// Mitsubishi GX Works2 project: TEAM_PLC   PLC: Q03UD

PROGRAM MAIN3
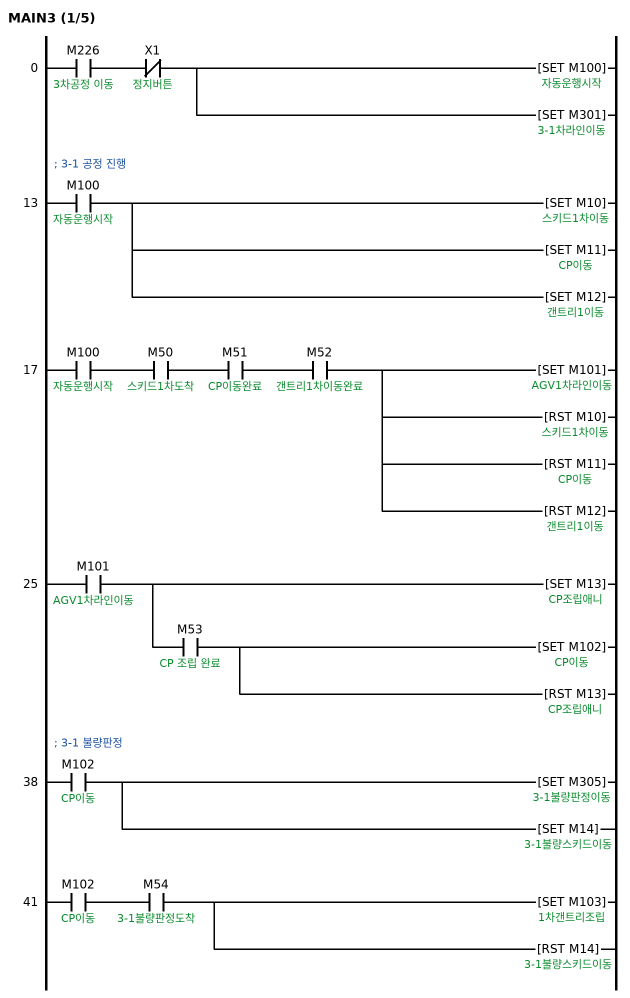
0     LD      M226  ; 3차공정 이동
      ANI     X1  ; 정지버튼
      SET     M100  ; 자동운행시작
      SET     M301  ; 3-1차라인이동
; 3-1 공정 진행
13    LD      M100  ; 자동운행시작
      SET     M10  ; 스키드1차이동
      SET     M11  ; CP이동
      SET     M12  ; 갠트리1이동
17    LD      M100  ; 자동운행시작
      AND     M50  ; 스키드1차도착
      AND     M51  ; CP이동완료
      AND     M52  ; 갠트리1차이동완료
      SET     M101  ; AGV1차라인이동
      RST     M10  ; 스키드1차이동
      RST     M11  ; CP이동
      RST     M12  ; 갠트리1이동
25    LD      M101  ; AGV1차라인이동
      SET     M13  ; CP조립애니
      AND     M53  ; CP 조립 완료
      SET     M102  ; CP이동
      RST     M13  ; CP조립애니
; 3-1 불량판정
38    LD      M102  ; CP이동
      SET     M305  ; 3-1불량판정이동
      SET     M14  ; 3-1불량스키드이동
41    LD      M102  ; CP이동
      AND     M54  ; 3-1불량판정도착
      SET     M103  ; 1차갠트리조립
      RST     M14  ; 3-1불량스키드이동
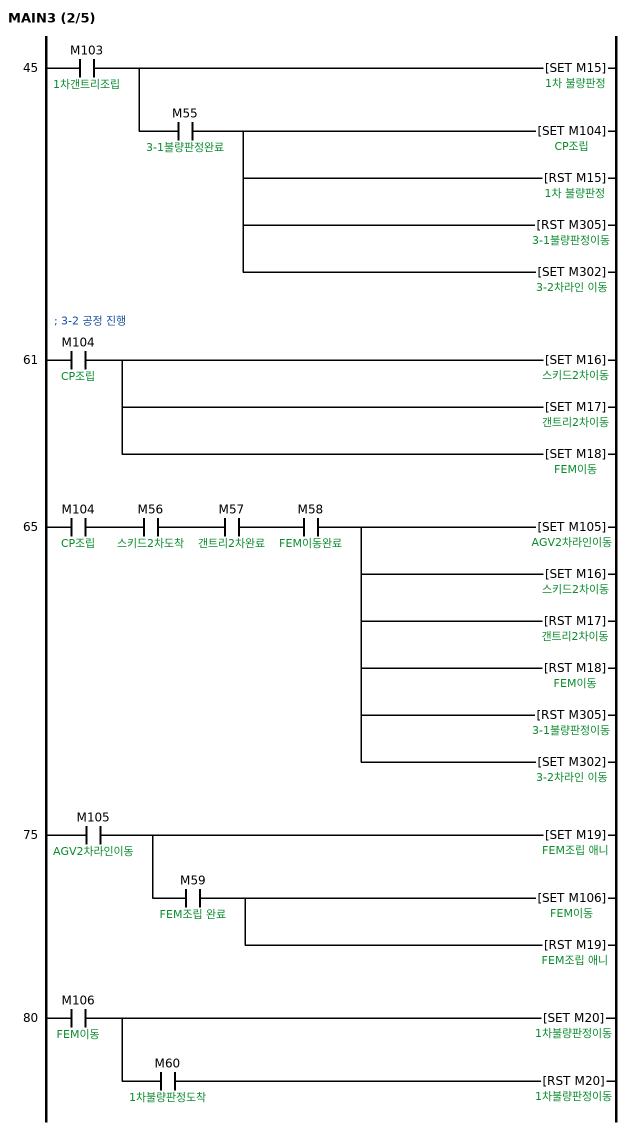
45    LD      M103  ; 1차갠트리조립
      SET     M15  ; 1차 불량판정
      AND     M55  ; 3-1불량판정완료
      SET     M104  ; CP조립
      RST     M15  ; 1차 불량판정
      RST     M305  ; 3-1불량판정이동
      SET     M302  ; 3-2차라인 이동
; 3-2 공정 진행
61    LD      M104  ; CP조립
      SET     M16  ; 스키드2차이동
      SET     M17  ; 갠트리2차이동
      SET     M18  ; FEM이동
65    LD      M104  ; CP조립
      AND     M56  ; 스키드2차도착
      AND     M57  ; 갠트리2차완료
      AND     M58  ; FEM이동완료
      SET     M105  ; AGV2차라인이동
      SET     M16  ; 스키드2차이동
      RST     M17  ; 갠트리2차이동
      RST     M18  ; FEM이동
      RST     M305  ; 3-1불량판정이동
      SET     M302  ; 3-2차라인 이동
75    LD      M105  ; AGV2차라인이동
      SET     M19  ; FEM조립 애니
      AND     M59  ; FEM조립 완료
      SET     M106  ; FEM이동
      RST     M19  ; FEM조립 애니
80    LD      M106  ; FEM이동
      SET     M20  ; 1차불량판정이동
      AND     M60  ; 1차불량판정도착
      RST     M20  ; 1차불량판정이동
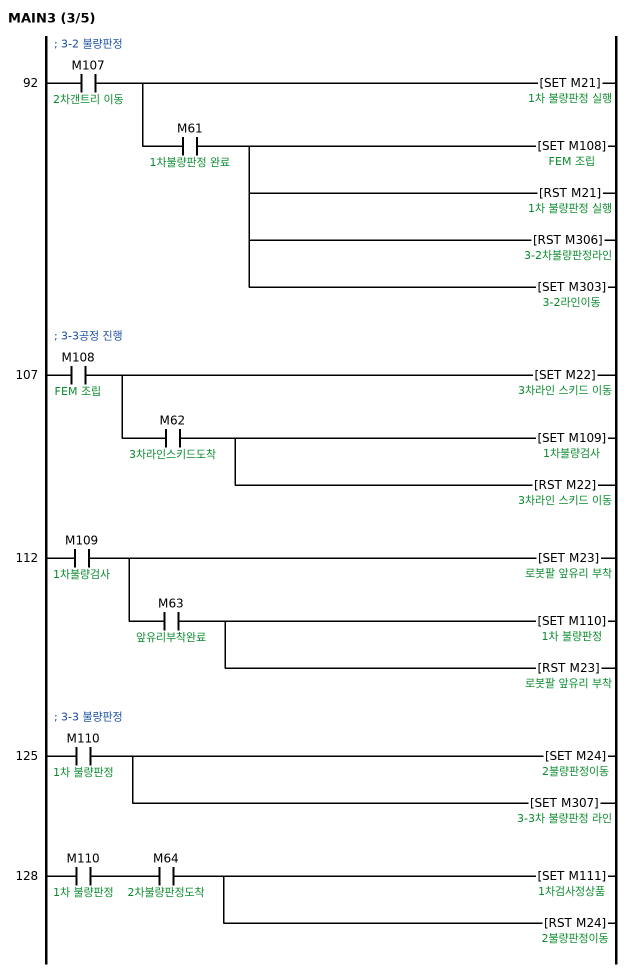
; 3-2 불량판정
92    LD      M107  ; 2차갠트리 이동
      SET     M21  ; 1차 불량판정 실행
      AND     M61  ; 1차불량판정 완료
      SET     M108  ; FEM 조립
      RST     M21  ; 1차 불량판정 실행
      RST     M306  ; 3-2차불량판정라인
      SET     M303  ; 3-2라인이동
; 3-3공정 진행
107   LD      M108  ; FEM 조립
      SET     M22  ; 3차라인 스키드 이동
      AND     M62  ; 3차라인스키드도착
      SET     M109  ; 1차불량검사
      RST     M22  ; 3차라인 스키드 이동
112   LD      M109  ; 1차불량검사
      SET     M23  ; 로봇팔 앞유리 부착
      AND     M63  ; 앞유리부착완료
      SET     M110  ; 1차 불량판정
      RST     M23  ; 로봇팔 앞유리 부착
; 3-3 불량판정
125   LD      M110  ; 1차 불량판정
      SET     M24  ; 2불량판정이동
      SET     M307  ; 3-3차 불량판정 라인
128   LD      M110  ; 1차 불량판정
      AND     M64  ; 2차불량판정도착
      SET     M111  ; 1차검사정상품
      RST     M24  ; 2불량판정이동
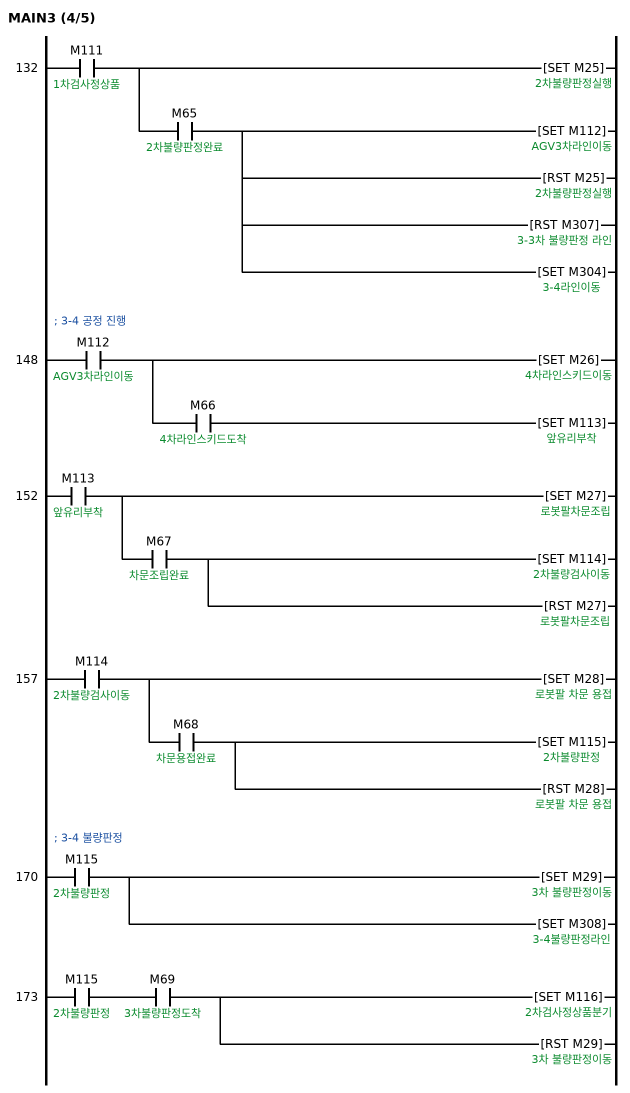
132   LD      M111  ; 1차검사정상품
      SET     M25  ; 2차불량판정실행
      AND     M65  ; 2차불량판정완료
      SET     M112  ; AGV3차라인이동
      RST     M25  ; 2차불량판정실행
      RST     M307  ; 3-3차 불량판정 라인
      SET     M304  ; 3-4라인이동
; 3-4 공정 진행
148   LD      M112  ; AGV3차라인이동
      SET     M26  ; 4차라인스키드이동
      AND     M66  ; 4차라인스키드도착
      SET     M113  ; 앞유리부착
152   LD      M113  ; 앞유리부착
      SET     M27  ; 로봇팔차문조립
      AND     M67  ; 차문조립완료
      SET     M114  ; 2차불량검사이동
      RST     M27  ; 로봇팔차문조립
157   LD      M114  ; 2차불량검사이동
      SET     M28  ; 로봇팔 차문 용접
      AND     M68  ; 차문용접완료
      SET     M115  ; 2차불량판정
      RST     M28  ; 로봇팔 차문 용접
; 3-4 불량판정
170   LD      M115  ; 2차불량판정
      SET     M29  ; 3차 불량판정이동
      SET     M308  ; 3-4불량판정라인
173   LD      M115  ; 2차불량판정
      AND     M69  ; 3차불량판정도착
      SET     M116  ; 2차검사정상품분기
      RST     M29  ; 3차 불량판정이동
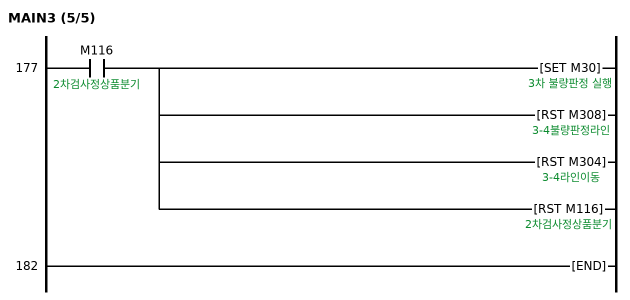
177   LD      M116  ; 2차검사정상품분기
      SET     M30  ; 3차 불량판정 실행
      RST     M308  ; 3-4불량판정라인
      RST     M304  ; 3-4라인이동
      RST     M116  ; 2차검사정상품분기
182   END
END_PROGRAM

PROGRAM MAIN1
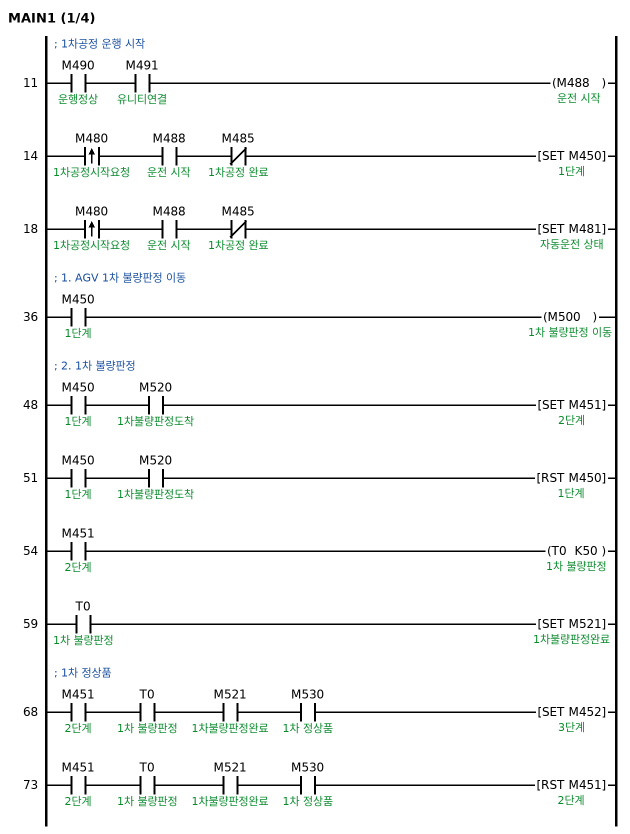
; 1차공정 운행 시작
11    LD      M490  ; 운행정상
      AND     M491  ; 유니티연결
      OUT     M488  ; 운전 시작
14    LDP     M480  ; 1차공정시작요청
      AND     M488  ; 운전 시작
      ANI     M485  ; 1차공정 완료
      SET     M450  ; 1단계
18    LDP     M480  ; 1차공정시작요청
      AND     M488  ; 운전 시작
      ANI     M485  ; 1차공정 완료
      SET     M481  ; 자동운전 상태
; 1. AGV 1차 불량판정 이동
36    LD      M450  ; 1단계
      OUT     M500  ; 1차 불량판정 이동
; 2. 1차 불량판정
48    LD      M450  ; 1단계
      AND     M520  ; 1차불량판정도착
      SET     M451  ; 2단계
51    LD      M450  ; 1단계
      AND     M520  ; 1차불량판정도착
      RST     M450  ; 1단계
54    LD      M451  ; 2단계
      OUT     T0 K50  ; 1차 불량판정
59    LD      T0  ; 1차 불량판정
      SET     M521  ; 1차불량판정완료
; 1차 정상품
68    LD      M451  ; 2단계
      AND     T0  ; 1차 불량판정
      AND     M521  ; 1차불량판정완료
      AND     M530  ; 1차 정상품
      SET     M452  ; 3단계
73    LD      M451  ; 2단계
      AND     T0  ; 1차 불량판정
      AND     M521  ; 1차불량판정완료
      AND     M530  ; 1차 정상품
      RST     M451  ; 2단계
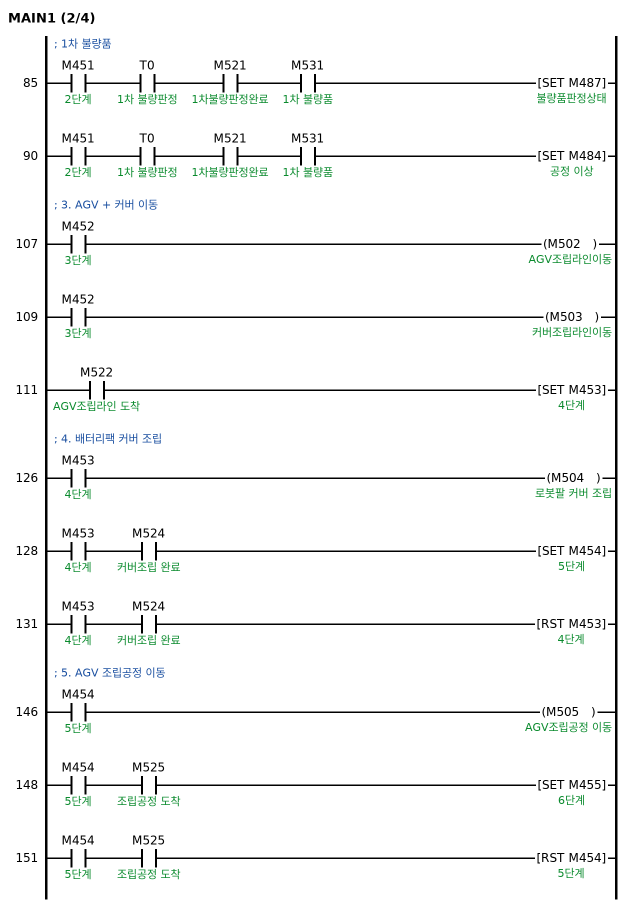
; 1차 불량품
85    LD      M451  ; 2단계
      AND     T0  ; 1차 불량판정
      AND     M521  ; 1차불량판정완료
      AND     M531  ; 1차 불량품
      SET     M487  ; 불량품판정상태
90    LD      M451  ; 2단계
      AND     T0  ; 1차 불량판정
      AND     M521  ; 1차불량판정완료
      AND     M531  ; 1차 불량품
      SET     M484  ; 공정 이상
; 3. AGV + 커버 이동
107   LD      M452  ; 3단계
      OUT     M502  ; AGV조립라인이동
109   LD      M452  ; 3단계
      OUT     M503  ; 커버조립라인이동
111   LD      M522  ; AGV조립라인 도착
      SET     M453  ; 4단계
; 4. 배터리팩 커버 조립
126   LD      M453  ; 4단계
      OUT     M504  ; 로봇팔 커버 조립
128   LD      M453  ; 4단계
      AND     M524  ; 커버조립 완료
      SET     M454  ; 5단계
131   LD      M453  ; 4단계
      AND     M524  ; 커버조립 완료
      RST     M453  ; 4단계
; 5. AGV 조립공정 이동
146   LD      M454  ; 5단계
      OUT     M505  ; AGV조립공정 이동
148   LD      M454  ; 5단계
      AND     M525  ; 조립공정 도착
      SET     M455  ; 6단계
151   LD      M454  ; 5단계
      AND     M525  ; 조립공정 도착
      RST     M454  ; 5단계
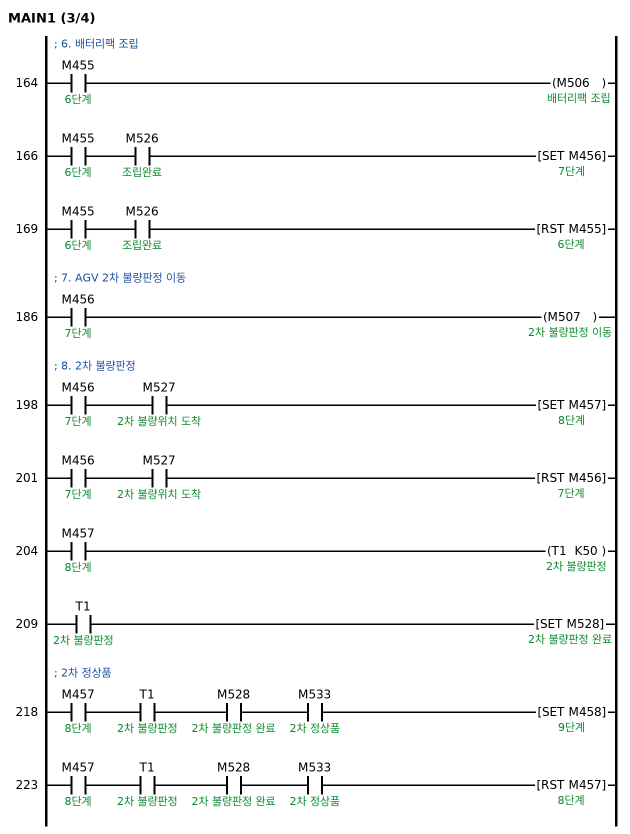
; 6. 배터리팩 조립
164   LD      M455  ; 6단계
      OUT     M506  ; 배터리팩 조립
166   LD      M455  ; 6단계
      AND     M526  ; 조립완료
      SET     M456  ; 7단계
169   LD      M455  ; 6단계
      AND     M526  ; 조립완료
      RST     M455  ; 6단계
; 7. AGV 2차 불량판정 이동
186   LD      M456  ; 7단계
      OUT     M507  ; 2차 불량판정 이동
; 8. 2차 불량판정
198   LD      M456  ; 7단계
      AND     M527  ; 2차 불량위치 도착
      SET     M457  ; 8단계
201   LD      M456  ; 7단계
      AND     M527  ; 2차 불량위치 도착
      RST     M456  ; 7단계
204   LD      M457  ; 8단계
      OUT     T1 K50  ; 2차 불량판정
209   LD      T1  ; 2차 불량판정
      SET     M528  ; 2차 불량판정 완료
; 2차 정상품
218   LD      M457  ; 8단계
      AND     T1  ; 2차 불량판정
      AND     M528  ; 2차 불량판정 완료
      AND     M533  ; 2차 정상품
      SET     M458  ; 9단계
223   LD      M457  ; 8단계
      AND     T1  ; 2차 불량판정
      AND     M528  ; 2차 불량판정 완료
      AND     M533  ; 2차 정상품
      RST     M457  ; 8단계
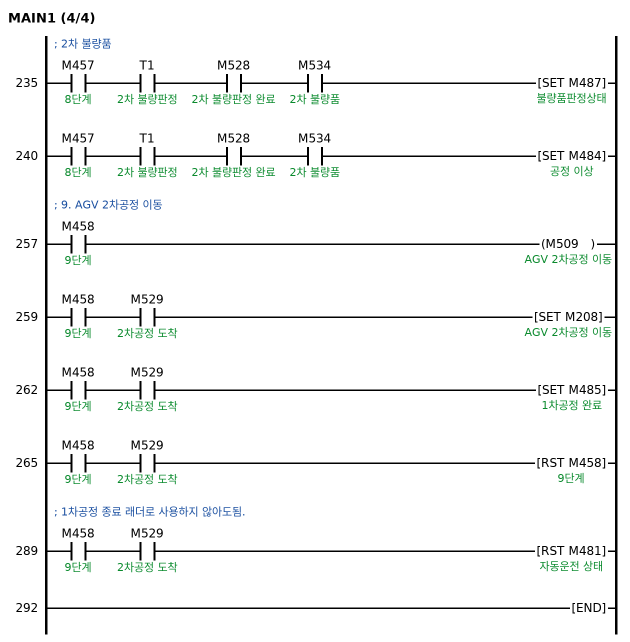
; 2차 불량품
235   LD      M457  ; 8단계
      AND     T1  ; 2차 불량판정
      AND     M528  ; 2차 불량판정 완료
      AND     M534  ; 2차 불량품
      SET     M487  ; 불량품판정상태
240   LD      M457  ; 8단계
      AND     T1  ; 2차 불량판정
      AND     M528  ; 2차 불량판정 완료
      AND     M534  ; 2차 불량품
      SET     M484  ; 공정 이상
; 9. AGV 2차공정 이동
257   LD      M458  ; 9단계
      OUT     M509  ; AGV 2차공정 이동
259   LD      M458  ; 9단계
      AND     M529  ; 2차공정 도착
      SET     M208  ; AGV 2차공정 이동
262   LD      M458  ; 9단계
      AND     M529  ; 2차공정 도착
      SET     M485  ; 1차공정 완료
265   LD      M458  ; 9단계
      AND     M529  ; 2차공정 도착
      RST     M458  ; 9단계
; 1차공정 종료 래더로 사용하지 않아도됨.
289   LD      M458  ; 9단계
      AND     M529  ; 2차공정 도착
      RST     M481  ; 자동운전 상태
292   END
END_PROGRAM

PROGRAM IOCHECK
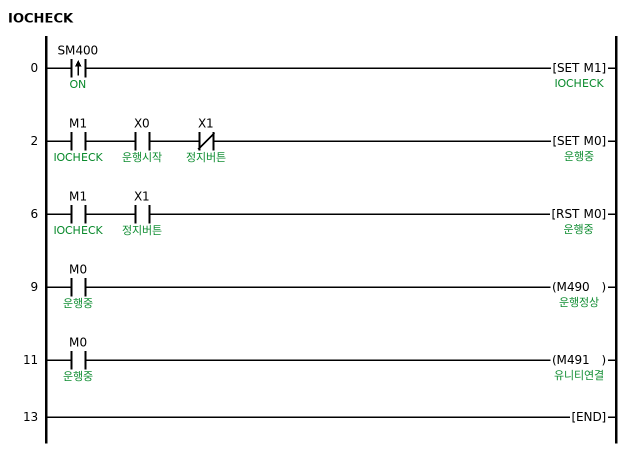
0     LDP     SM400  ; ON
      SET     M1  ; IOCHECK
2     LD      M1  ; IOCHECK
      AND     X0  ; 운행시작
      ANI     X1  ; 정지버튼
      SET     M0  ; 운행중
6     LD      M1  ; IOCHECK
      AND     X1  ; 정지버튼
      RST     M0  ; 운행중
9     LD      M0  ; 운행중
      OUT     M490  ; 운행정상
11    LD      M0  ; 운행중
      OUT     M491  ; 유니티연결
13    END
END_PROGRAM

PROGRAM MAIN2
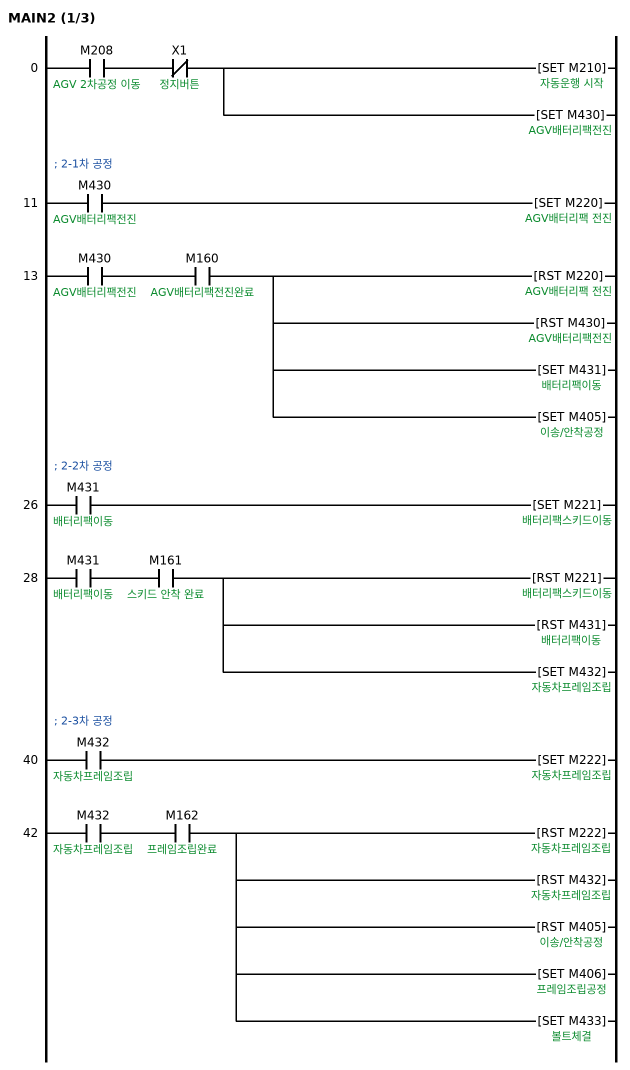
0     LD      M208  ; AGV 2차공정 이동
      ANI     X1  ; 정지버튼
      SET     M210  ; 자동운행 시작
      SET     M430  ; AGV배터리팩전진
; 2-1차 공정
11    LD      M430  ; AGV배터리팩전진
      SET     M220  ; AGV배터리팩 전진
13    LD      M430  ; AGV배터리팩전진
      AND     M160  ; AGV배터리팩전진완료
      RST     M220  ; AGV배터리팩 전진
      RST     M430  ; AGV배터리팩전진
      SET     M431  ; 배터리팩이동
      SET     M405  ; 이송/안착공정
; 2-2차 공정
26    LD      M431  ; 배터리팩이동
      SET     M221  ; 배터리팩스키드이동
28    LD      M431  ; 배터리팩이동
      AND     M161  ; 스키드 안착 완료
      RST     M221  ; 배터리팩스키드이동
      RST     M431  ; 배터리팩이동
      SET     M432  ; 자동차프레임조립
; 2-3차 공정
40    LD      M432  ; 자동차프레임조립
      SET     M222  ; 자동차프레임조립
42    LD      M432  ; 자동차프레임조립
      AND     M162  ; 프레임조립완료
      RST     M222  ; 자동차프레임조립
      RST     M432  ; 자동차프레임조립
      RST     M405  ; 이송/안착공정
      SET     M406  ; 프레임조립공정
      SET     M433  ; 볼트체결
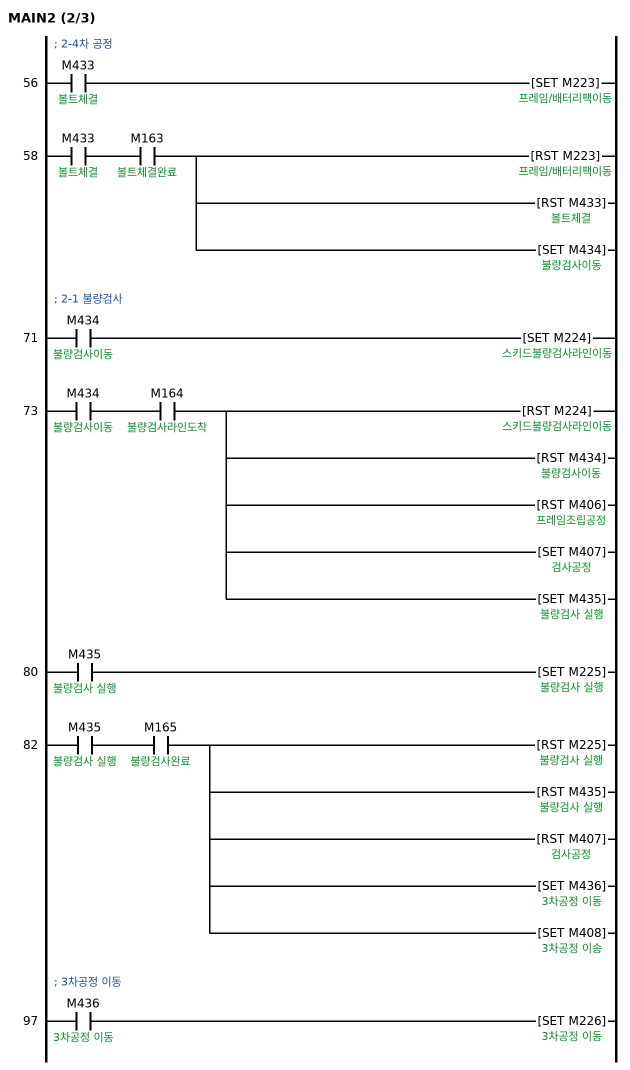
; 2-4차 공정
56    LD      M433  ; 볼트체결
      SET     M223  ; 프레임/배터리팩이동
58    LD      M433  ; 볼트체결
      AND     M163  ; 볼트체결완료
      RST     M223  ; 프레임/배터리팩이동
      RST     M433  ; 볼트체결
      SET     M434  ; 불량검사이동
; 2-1 불량검사
71    LD      M434  ; 불량검사이동
      SET     M224  ; 스키드불량검사라인이동
73    LD      M434  ; 불량검사이동
      AND     M164  ; 불량검사라인도착
      RST     M224  ; 스키드불량검사라인이동
      RST     M434  ; 불량검사이동
      RST     M406  ; 프레임조립공정
      SET     M407  ; 검사공정
      SET     M435  ; 불량검사 실행
80    LD      M435  ; 불량검사 실행
      SET     M225  ; 불량검사 실행
82    LD      M435  ; 불량검사 실행
      AND     M165  ; 불량검사완료
      RST     M225  ; 불량검사 실행
      RST     M435  ; 불량검사 실행
      RST     M407  ; 검사공정
      SET     M436  ; 3차공정 이동
      SET     M408  ; 3차공정 이송
; 3차공정 이동
97    LD      M436  ; 3차공정 이동
      SET     M226  ; 3차공정 이동
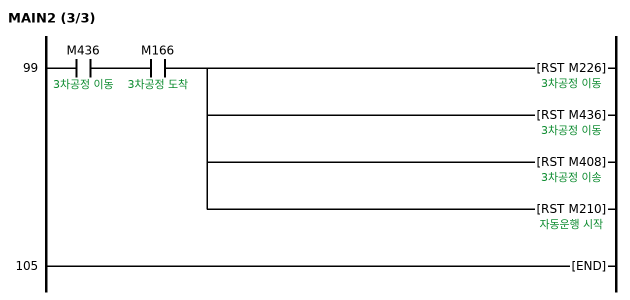
99    LD      M436  ; 3차공정 이동
      AND     M166  ; 3차공정 도착
      RST     M226  ; 3차공정 이동
      RST     M436  ; 3차공정 이동
      RST     M408  ; 3차공정 이송
      RST     M210  ; 자동운행 시작
105   END
END_PROGRAM

PROGRAM MAIN1-1
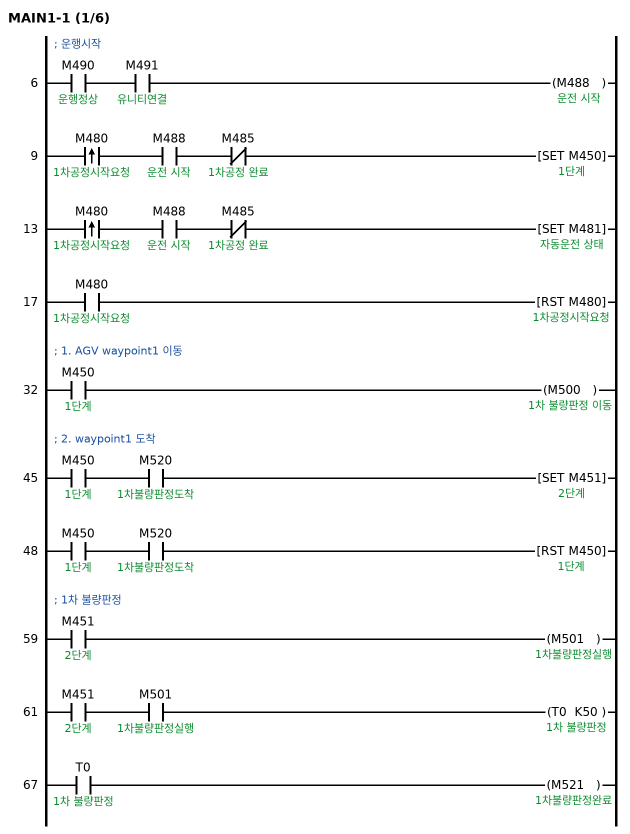
; 운행시작
6     LD      M490  ; 운행정상
      AND     M491  ; 유니티연결
      OUT     M488  ; 운전 시작
9     LDP     M480  ; 1차공정시작요청
      AND     M488  ; 운전 시작
      ANI     M485  ; 1차공정 완료
      SET     M450  ; 1단계
13    LDP     M480  ; 1차공정시작요청
      AND     M488  ; 운전 시작
      ANI     M485  ; 1차공정 완료
      SET     M481  ; 자동운전 상태
17    LD      M480  ; 1차공정시작요청
      RST     M480  ; 1차공정시작요청
; 1. AGV waypoint1 이동
32    LD      M450  ; 1단계
      OUT     M500  ; 1차 불량판정 이동
; 2. waypoint1 도착
45    LD      M450  ; 1단계
      AND     M520  ; 1차불량판정도착
      SET     M451  ; 2단계
48    LD      M450  ; 1단계
      AND     M520  ; 1차불량판정도착
      RST     M450  ; 1단계
; 1차 불량판정
59    LD      M451  ; 2단계
      OUT     M501  ; 1차불량판정실행
61    LD      M451  ; 2단계
      AND     M501  ; 1차불량판정실행
      OUT     T0 K50  ; 1차 불량판정
67    LD      T0  ; 1차 불량판정
      OUT     M521  ; 1차불량판정완료
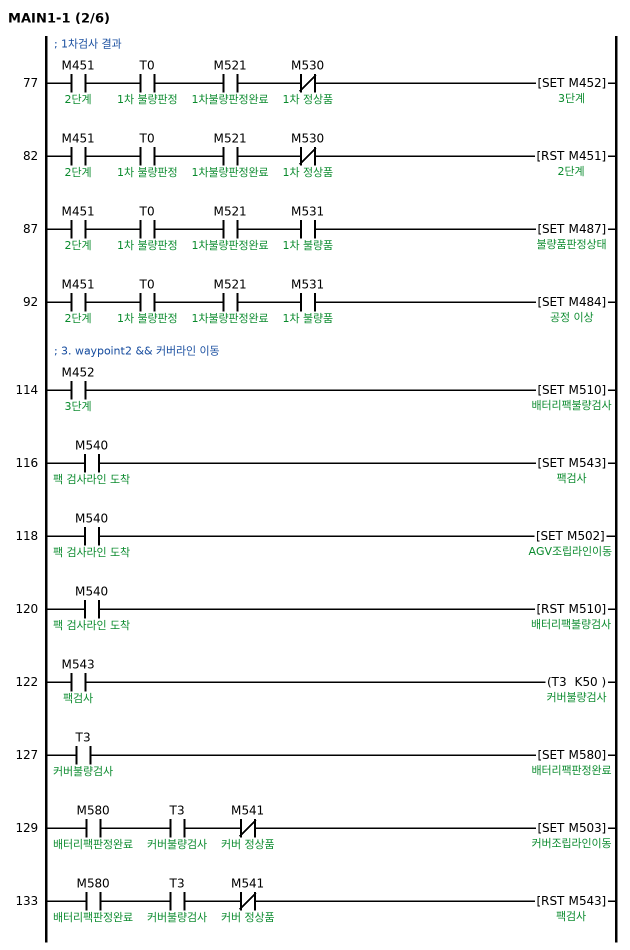
; 1차검사 결과
77    LD      M451  ; 2단계
      AND     T0  ; 1차 불량판정
      AND     M521  ; 1차불량판정완료
      ANI     M530  ; 1차 정상품
      SET     M452  ; 3단계
82    LD      M451  ; 2단계
      AND     T0  ; 1차 불량판정
      AND     M521  ; 1차불량판정완료
      ANI     M530  ; 1차 정상품
      RST     M451  ; 2단계
87    LD      M451  ; 2단계
      AND     T0  ; 1차 불량판정
      AND     M521  ; 1차불량판정완료
      AND     M531  ; 1차 불량품
      SET     M487  ; 불량품판정상태
92    LD      M451  ; 2단계
      AND     T0  ; 1차 불량판정
      AND     M521  ; 1차불량판정완료
      AND     M531  ; 1차 불량품
      SET     M484  ; 공정 이상
; 3. waypoint2 && 커버라인 이동
114   LD      M452  ; 3단계
      SET     M510  ; 배터리팩불량검사
116   LD      M540  ; 팩 검사라인 도착
      SET     M543  ; 팩검사
118   LD      M540  ; 팩 검사라인 도착
      SET     M502  ; AGV조립라인이동
120   LD      M540  ; 팩 검사라인 도착
      RST     M510  ; 배터리팩불량검사
122   LD      M543  ; 팩검사
      OUT     T3 K50  ; 커버불량검사
127   LD      T3  ; 커버불량검사
      SET     M580  ; 배터리팩판정완료
129   LD      M580  ; 배터리팩판정완료
      AND     T3  ; 커버불량검사
      ANI     M541  ; 커버 정상품
      SET     M503  ; 커버조립라인이동
133   LD      M580  ; 배터리팩판정완료
      AND     T3  ; 커버불량검사
      ANI     M541  ; 커버 정상품
      RST     M543  ; 팩검사
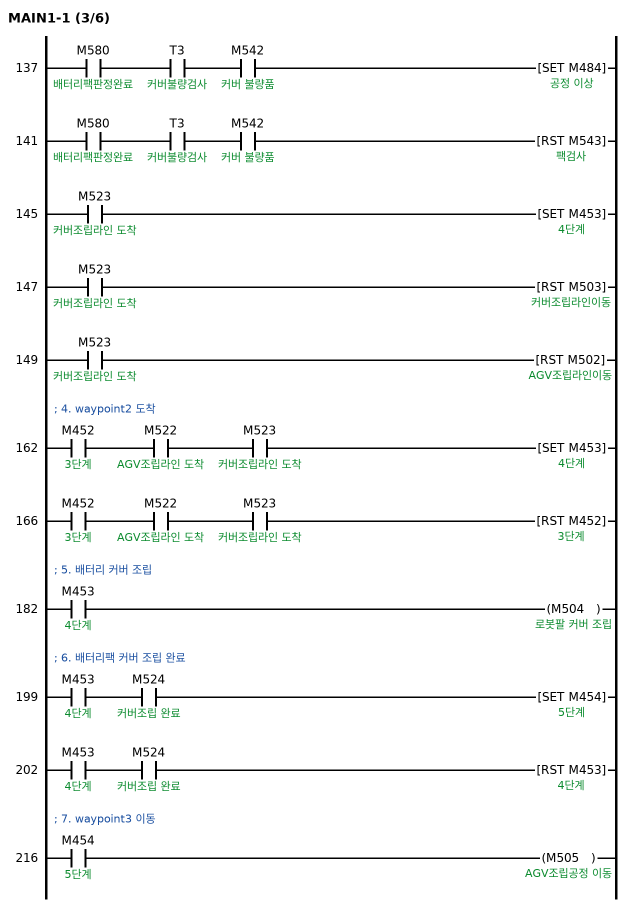
137   LD      M580  ; 배터리팩판정완료
      AND     T3  ; 커버불량검사
      AND     M542  ; 커버 불량품
      SET     M484  ; 공정 이상
141   LD      M580  ; 배터리팩판정완료
      AND     T3  ; 커버불량검사
      AND     M542  ; 커버 불량품
      RST     M543  ; 팩검사
145   LD      M523  ; 커버조립라인 도착
      SET     M453  ; 4단계
147   LD      M523  ; 커버조립라인 도착
      RST     M503  ; 커버조립라인이동
149   LD      M523  ; 커버조립라인 도착
      RST     M502  ; AGV조립라인이동
; 4. waypoint2 도착
162   LD      M452  ; 3단계
      AND     M522  ; AGV조립라인 도착
      AND     M523  ; 커버조립라인 도착
      SET     M453  ; 4단계
166   LD      M452  ; 3단계
      AND     M522  ; AGV조립라인 도착
      AND     M523  ; 커버조립라인 도착
      RST     M452  ; 3단계
; 5. 배터리 커버 조립
182   LD      M453  ; 4단계
      OUT     M504  ; 로봇팔 커버 조립
; 6. 배터리팩 커버 조립 완료
199   LD      M453  ; 4단계
      AND     M524  ; 커버조립 완료
      SET     M454  ; 5단계
202   LD      M453  ; 4단계
      AND     M524  ; 커버조립 완료
      RST     M453  ; 4단계
; 7. waypoint3 이동
216   LD      M454  ; 5단계
      OUT     M505  ; AGV조립공정 이동
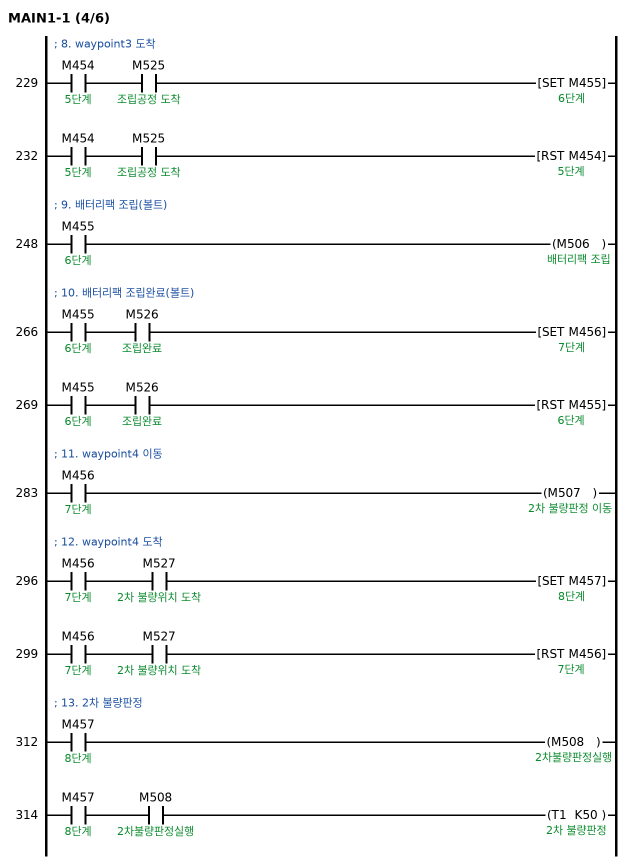
; 8. waypoint3 도착
229   LD      M454  ; 5단계
      AND     M525  ; 조립공정 도착
      SET     M455  ; 6단계
232   LD      M454  ; 5단계
      AND     M525  ; 조립공정 도착
      RST     M454  ; 5단계
; 9. 배터리팩 조립(볼트)
248   LD      M455  ; 6단계
      OUT     M506  ; 배터리팩 조립
; 10. 배터리팩 조립완료(볼트)
266   LD      M455  ; 6단계
      AND     M526  ; 조립완료
      SET     M456  ; 7단계
269   LD      M455  ; 6단계
      AND     M526  ; 조립완료
      RST     M455  ; 6단계
; 11. waypoint4 이동
283   LD      M456  ; 7단계
      OUT     M507  ; 2차 불량판정 이동
; 12. waypoint4 도착
296   LD      M456  ; 7단계
      AND     M527  ; 2차 불량위치 도착
      SET     M457  ; 8단계
299   LD      M456  ; 7단계
      AND     M527  ; 2차 불량위치 도착
      RST     M456  ; 7단계
; 13. 2차 불량판정
312   LD      M457  ; 8단계
      OUT     M508  ; 2차불량판정실행
314   LD      M457  ; 8단계
      AND     M508  ; 2차불량판정실행
      OUT     T1 K50  ; 2차 불량판정
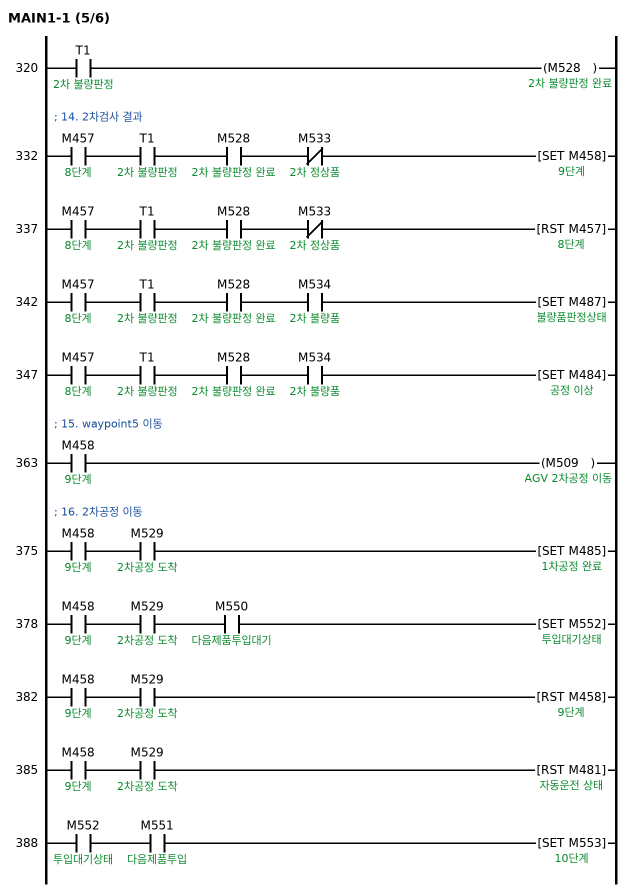
320   LD      T1  ; 2차 불량판정
      OUT     M528  ; 2차 불량판정 완료
; 14. 2차검사 결과
332   LD      M457  ; 8단계
      AND     T1  ; 2차 불량판정
      AND     M528  ; 2차 불량판정 완료
      ANI     M533  ; 2차 정상품
      SET     M458  ; 9단계
337   LD      M457  ; 8단계
      AND     T1  ; 2차 불량판정
      AND     M528  ; 2차 불량판정 완료
      ANI     M533  ; 2차 정상품
      RST     M457  ; 8단계
342   LD      M457  ; 8단계
      AND     T1  ; 2차 불량판정
      AND     M528  ; 2차 불량판정 완료
      AND     M534  ; 2차 불량품
      SET     M487  ; 불량품판정상태
347   LD      M457  ; 8단계
      AND     T1  ; 2차 불량판정
      AND     M528  ; 2차 불량판정 완료
      AND     M534  ; 2차 불량품
      SET     M484  ; 공정 이상
; 15. waypoint5 이동
363   LD      M458  ; 9단계
      OUT     M509  ; AGV 2차공정 이동
; 16. 2차공정 이동
375   LD      M458  ; 9단계
      AND     M529  ; 2차공정 도착
      SET     M485  ; 1차공정 완료
378   LD      M458  ; 9단계
      AND     M529  ; 2차공정 도착
      AND     M550  ; 다음제품투입대기
      SET     M552  ; 투입대기상태
382   LD      M458  ; 9단계
      AND     M529  ; 2차공정 도착
      RST     M458  ; 9단계
385   LD      M458  ; 9단계
      AND     M529  ; 2차공정 도착
      RST     M481  ; 자동운전 상태
388   LD      M552  ; 투입대기상태
      AND     M551  ; 다음제품투입
      SET     M553  ; 10단계
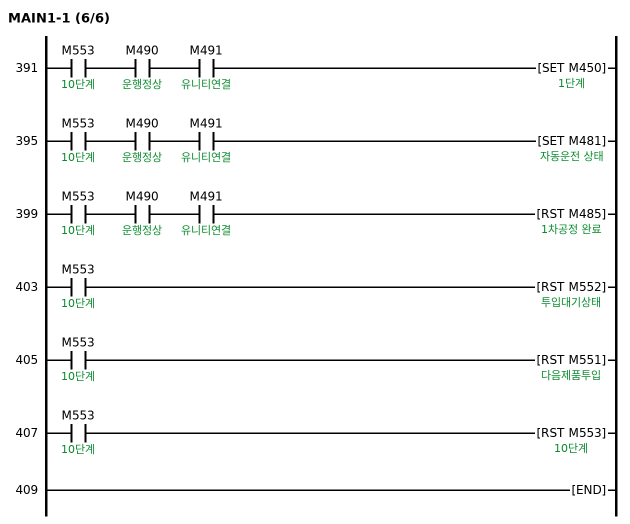
391   LD      M553  ; 10단계
      AND     M490  ; 운행정상
      AND     M491  ; 유니티연결
      SET     M450  ; 1단계
395   LD      M553  ; 10단계
      AND     M490  ; 운행정상
      AND     M491  ; 유니티연결
      SET     M481  ; 자동운전 상태
399   LD      M553  ; 10단계
      AND     M490  ; 운행정상
      AND     M491  ; 유니티연결
      RST     M485  ; 1차공정 완료
403   LD      M553  ; 10단계
      RST     M552  ; 투입대기상태
405   LD      M553  ; 10단계
      RST     M551  ; 다음제품투입
407   LD      M553  ; 10단계
      RST     M553  ; 10단계
409   END
END_PROGRAM

PROGRAM MAIN3-1
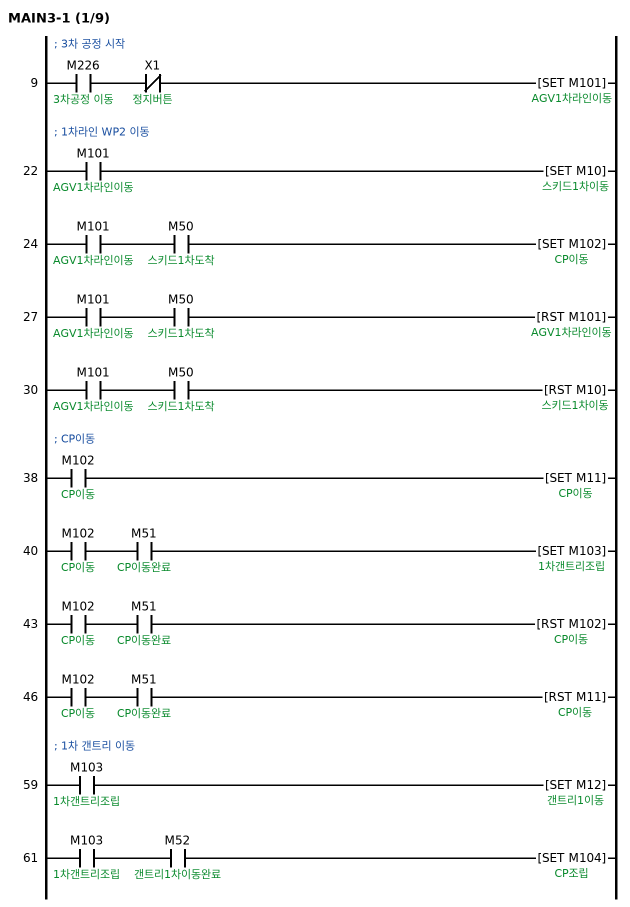
; 3차 공정 시작
9     LD      M226  ; 3차공정 이동
      ANI     X1  ; 정지버튼
      SET     M101  ; AGV1차라인이동
; 1차라인 WP2 이동
22    LD      M101  ; AGV1차라인이동
      SET     M10  ; 스키드1차이동
24    LD      M101  ; AGV1차라인이동
      AND     M50  ; 스키드1차도착
      SET     M102  ; CP이동
27    LD      M101  ; AGV1차라인이동
      AND     M50  ; 스키드1차도착
      RST     M101  ; AGV1차라인이동
30    LD      M101  ; AGV1차라인이동
      AND     M50  ; 스키드1차도착
      RST     M10  ; 스키드1차이동
; CP이동
38    LD      M102  ; CP이동
      SET     M11  ; CP이동
40    LD      M102  ; CP이동
      AND     M51  ; CP이동완료
      SET     M103  ; 1차갠트리조립
43    LD      M102  ; CP이동
      AND     M51  ; CP이동완료
      RST     M102  ; CP이동
46    LD      M102  ; CP이동
      AND     M51  ; CP이동완료
      RST     M11  ; CP이동
; 1차 갠트리 이동
59    LD      M103  ; 1차갠트리조립
      SET     M12  ; 갠트리1이동
61    LD      M103  ; 1차갠트리조립
      AND     M52  ; 갠트리1차이동완료
      SET     M104  ; CP조립
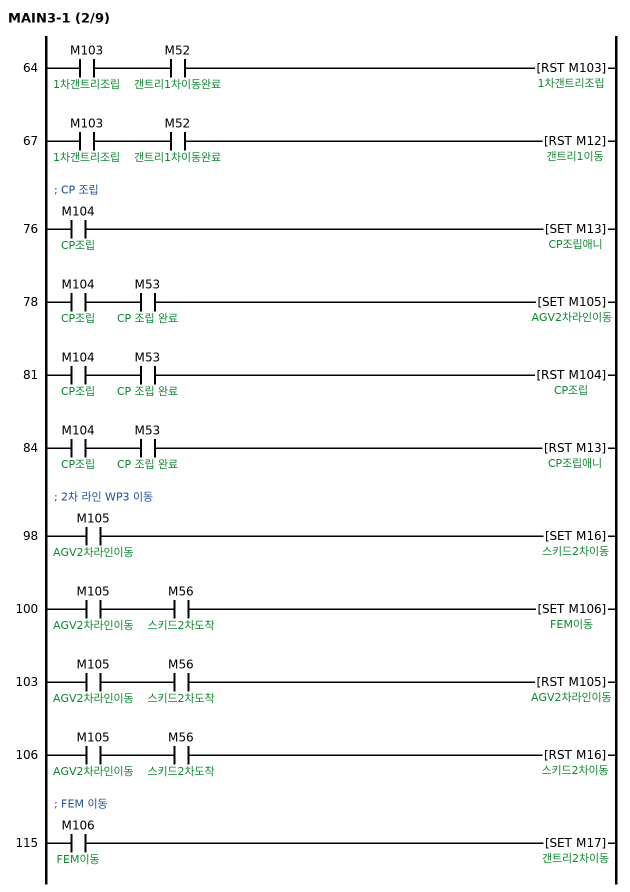
64    LD      M103  ; 1차갠트리조립
      AND     M52  ; 갠트리1차이동완료
      RST     M103  ; 1차갠트리조립
67    LD      M103  ; 1차갠트리조립
      AND     M52  ; 갠트리1차이동완료
      RST     M12  ; 갠트리1이동
; CP 조립
76    LD      M104  ; CP조립
      SET     M13  ; CP조립애니
78    LD      M104  ; CP조립
      AND     M53  ; CP 조립 완료
      SET     M105  ; AGV2차라인이동
81    LD      M104  ; CP조립
      AND     M53  ; CP 조립 완료
      RST     M104  ; CP조립
84    LD      M104  ; CP조립
      AND     M53  ; CP 조립 완료
      RST     M13  ; CP조립애니
; 2차 라인 WP3 이동
98    LD      M105  ; AGV2차라인이동
      SET     M16  ; 스키드2차이동
100   LD      M105  ; AGV2차라인이동
      AND     M56  ; 스키드2차도착
      SET     M106  ; FEM이동
103   LD      M105  ; AGV2차라인이동
      AND     M56  ; 스키드2차도착
      RST     M105  ; AGV2차라인이동
106   LD      M105  ; AGV2차라인이동
      AND     M56  ; 스키드2차도착
      RST     M16  ; 스키드2차이동
; FEM 이동
115   LD      M106  ; FEM이동
      SET     M17  ; 갠트리2차이동
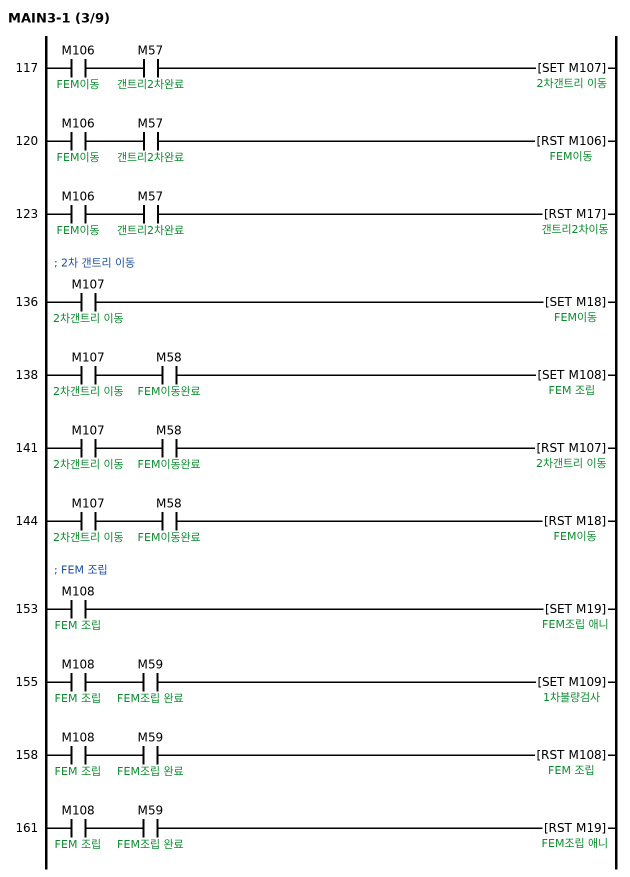
117   LD      M106  ; FEM이동
      AND     M57  ; 갠트리2차완료
      SET     M107  ; 2차갠트리 이동
120   LD      M106  ; FEM이동
      AND     M57  ; 갠트리2차완료
      RST     M106  ; FEM이동
123   LD      M106  ; FEM이동
      AND     M57  ; 갠트리2차완료
      RST     M17  ; 갠트리2차이동
; 2차 갠트리 이동
136   LD      M107  ; 2차갠트리 이동
      SET     M18  ; FEM이동
138   LD      M107  ; 2차갠트리 이동
      AND     M58  ; FEM이동완료
      SET     M108  ; FEM 조립
141   LD      M107  ; 2차갠트리 이동
      AND     M58  ; FEM이동완료
      RST     M107  ; 2차갠트리 이동
144   LD      M107  ; 2차갠트리 이동
      AND     M58  ; FEM이동완료
      RST     M18  ; FEM이동
; FEM 조립
153   LD      M108  ; FEM 조립
      SET     M19  ; FEM조립 애니
155   LD      M108  ; FEM 조립
      AND     M59  ; FEM조립 완료
      SET     M109  ; 1차불량검사
158   LD      M108  ; FEM 조립
      AND     M59  ; FEM조립 완료
      RST     M108  ; FEM 조립
161   LD      M108  ; FEM 조립
      AND     M59  ; FEM조립 완료
      RST     M19  ; FEM조립 애니
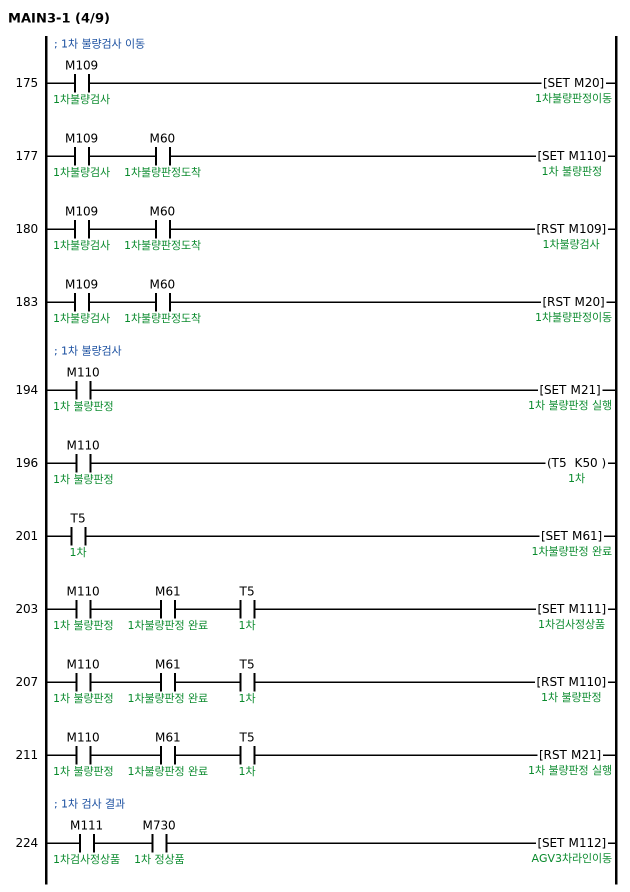
; 1차 불량검사 이동
175   LD      M109  ; 1차불량검사
      SET     M20  ; 1차불량판정이동
177   LD      M109  ; 1차불량검사
      AND     M60  ; 1차불량판정도착
      SET     M110  ; 1차 불량판정
180   LD      M109  ; 1차불량검사
      AND     M60  ; 1차불량판정도착
      RST     M109  ; 1차불량검사
183   LD      M109  ; 1차불량검사
      AND     M60  ; 1차불량판정도착
      RST     M20  ; 1차불량판정이동
; 1차 불량검사
194   LD      M110  ; 1차 불량판정
      SET     M21  ; 1차 불량판정 실행
196   LD      M110  ; 1차 불량판정
      OUT     T5 K50  ; 1차
201   LD      T5  ; 1차
      SET     M61  ; 1차불량판정 완료
203   LD      M110  ; 1차 불량판정
      AND     M61  ; 1차불량판정 완료
      AND     T5  ; 1차
      SET     M111  ; 1차검사정상품
207   LD      M110  ; 1차 불량판정
      AND     M61  ; 1차불량판정 완료
      AND     T5  ; 1차
      RST     M110  ; 1차 불량판정
211   LD      M110  ; 1차 불량판정
      AND     M61  ; 1차불량판정 완료
      AND     T5  ; 1차
      RST     M21  ; 1차 불량판정 실행
; 1차 검사 결과
224   LD      M111  ; 1차검사정상품
      AND     M730  ; 1차 정상품
      SET     M112  ; AGV3차라인이동
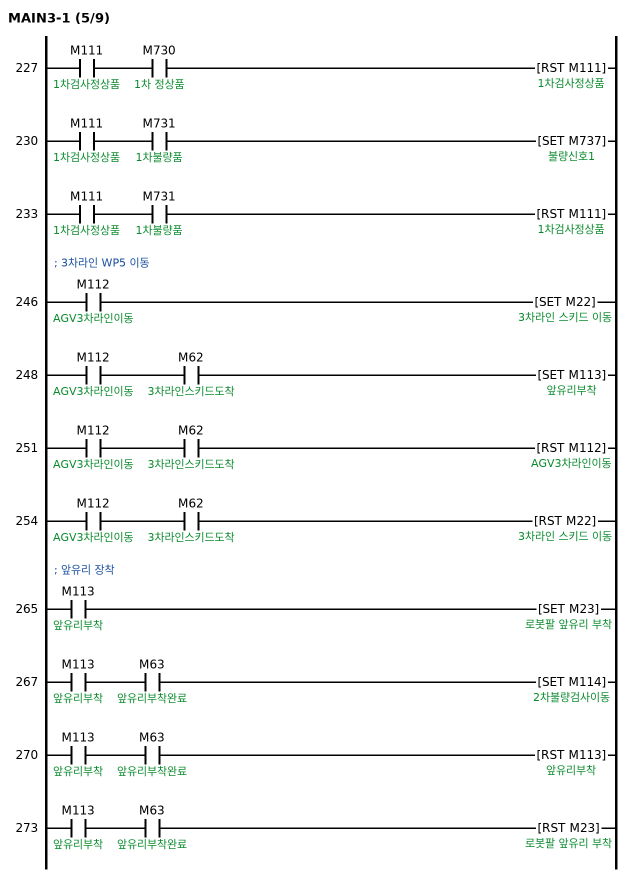
227   LD      M111  ; 1차검사정상품
      AND     M730  ; 1차 정상품
      RST     M111  ; 1차검사정상품
230   LD      M111  ; 1차검사정상품
      AND     M731  ; 1차불량품
      SET     M737  ; 불량신호1
233   LD      M111  ; 1차검사정상품
      AND     M731  ; 1차불량품
      RST     M111  ; 1차검사정상품
; 3차라인 WP5 이동
246   LD      M112  ; AGV3차라인이동
      SET     M22  ; 3차라인 스키드 이동
248   LD      M112  ; AGV3차라인이동
      AND     M62  ; 3차라인스키드도착
      SET     M113  ; 앞유리부착
251   LD      M112  ; AGV3차라인이동
      AND     M62  ; 3차라인스키드도착
      RST     M112  ; AGV3차라인이동
254   LD      M112  ; AGV3차라인이동
      AND     M62  ; 3차라인스키드도착
      RST     M22  ; 3차라인 스키드 이동
; 앞유리 장착
265   LD      M113  ; 앞유리부착
      SET     M23  ; 로봇팔 앞유리 부착
267   LD      M113  ; 앞유리부착
      AND     M63  ; 앞유리부착완료
      SET     M114  ; 2차불량검사이동
270   LD      M113  ; 앞유리부착
      AND     M63  ; 앞유리부착완료
      RST     M113  ; 앞유리부착
273   LD      M113  ; 앞유리부착
      AND     M63  ; 앞유리부착완료
      RST     M23  ; 로봇팔 앞유리 부착
